Yaskawa INFORM job: UTEST.JBI

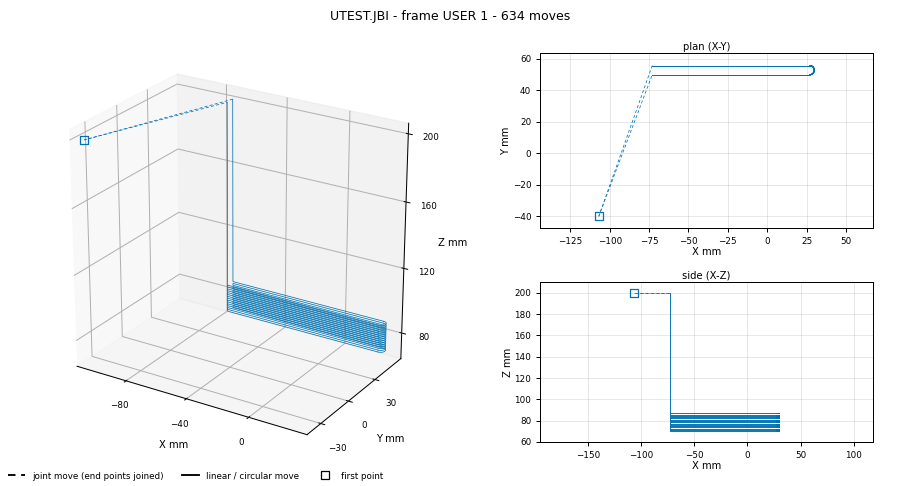
[picture p0: tool path of UTEST.JBI in frame USER 1, 634 of 649 moves have a stored position in this frame; points joined in program order, loops and branches not executed]
/JOB
//NAME UTEST
//POS
///NPOS 649,0,0,0,0,0
///USER 1
///TOOL 1
///POSTYPE USER
///RECTAN
///RCONF 1,0,0,0,0,0,0,0,0,0,0,0,0,0,0,0,0,0,0,0,0,0,0,0
C00000=-107.000,-40.000,200.000,0.0000,0.0000,-150.0000
C00001=-73.000,50.000,200.000,0.0000,0.0000,-150.0000
C00002=-73.000,50.000,70.000,0.0000,0.0000,-150.0000
C00003=-68.000,50.000,70.000,0.0000,0.0000,-150.0000
C00004=-63.000,50.000,70.000,0.0000,0.0000,-150.0000
C00005=-58.000,50.000,70.000,0.0000,0.0000,-150.0000
C00006=-53.000,50.000,70.000,0.0000,0.0000,-150.0000
C00007=-48.000,50.000,70.000,0.0000,0.0000,-150.0000
C00008=-43.000,50.000,70.000,0.0000,0.0000,-150.0000
C00009=-38.000,50.000,70.000,0.0000,0.0000,-150.0000
C00010=-33.000,50.000,70.000,0.0000,0.0000,-150.0000
C00011=-28.000,50.000,70.000,0.0000,0.0000,-150.0000
C00012=-23.000,50.000,70.000,0.0000,0.0000,-150.0000
C00013=-18.000,50.000,70.000,0.0000,0.0000,-150.0000
C00014=-13.000,50.000,70.000,0.0000,0.0000,-150.0000
C00015=-8.000,50.000,70.000,0.0000,0.0000,-150.0000
C00016=-3.000,50.000,70.000,0.0000,0.0000,-150.0000
C00017=2.000,50.000,70.000,0.0000,0.0000,-150.0000
C00018=7.000,50.000,70.000,0.0000,0.0000,-150.0000
C00019=12.000,50.000,70.000,0.0000,0.0000,-150.0000
C00020=17.000,50.000,70.000,0.0000,0.0000,-150.0000
C00021=22.000,50.000,70.000,0.0000,0.0000,-150.0000
C00022=27.000,50.000,70.000,0.0000,0.0000,-150.0000
C00023=29.915,52.915,70.000,0.0000,0.0000,-150.0000
C00024=27.000,55.829,70.000,0.0000,0.0000,-150.0000
C00025=22.000,55.829,70.000,0.0000,0.0000,-150.0000
C00026=17.000,55.829,70.000,0.0000,0.0000,-150.0000
C00027=12.000,55.829,70.000,0.0000,0.0000,-150.0000
C00028=7.000,55.829,70.000,0.0000,0.0000,-150.0000
C00029=2.000,55.829,70.000,0.0000,0.0000,-150.0000
C00030=-3.000,55.829,70.000,0.0000,0.0000,-150.0000
C00031=-8.000,55.829,70.000,0.0000,0.0000,-150.0000
C00032=-13.000,55.829,70.000,0.0000,0.0000,-150.0000
C00033=-18.000,55.829,70.000,0.0000,0.0000,-150.0000
C00034=-23.000,55.829,70.000,0.0000,0.0000,-150.0000
C00035=-28.000,55.829,70.000,0.0000,0.0000,-150.0000
C00036=-33.000,55.829,70.000,0.0000,0.0000,-150.0000
C00037=-38.000,55.829,70.000,0.0000,0.0000,-150.0000
C00038=-43.000,55.829,70.000,0.0000,0.0000,-150.0000
C00039=-48.000,55.829,70.000,0.0000,0.0000,-150.0000
C00040=-53.000,55.829,70.000,0.0000,0.0000,-150.0000
C00041=-58.000,55.829,70.000,0.0000,0.0000,-150.0000
C00042=-63.000,55.829,70.000,0.0000,0.0000,-150.0000
C00043=-68.000,55.829,70.000,0.0000,0.0000,-150.0000
C00044=-73.000,55.829,70.000,0.0000,0.0000,-150.0000
C00045=-73.000,55.829,71.200,0.0000,0.0000,-150.0000
C00046=-68.000,55.829,71.200,0.0000,0.0000,-150.0000
C00047=-63.000,55.829,71.200,0.0000,0.0000,-150.0000
C00048=-58.000,55.829,71.200,0.0000,0.0000,-150.0000
C00049=-53.000,55.829,71.200,0.0000,0.0000,-150.0000
C00050=-48.000,55.829,71.200,0.0000,0.0000,-150.0000
C00051=-43.000,55.829,71.200,0.0000,0.0000,-150.0000
C00052=-38.000,55.829,71.200,0.0000,0.0000,-150.0000
C00053=-33.000,55.829,71.200,0.0000,0.0000,-150.0000
C00054=-28.000,55.829,71.200,0.0000,0.0000,-150.0000
C00055=-23.000,55.829,71.200,0.0000,0.0000,-150.0000
C00056=-18.000,55.829,71.200,0.0000,0.0000,-150.0000
C00057=-13.000,55.829,71.200,0.0000,0.0000,-150.0000
C00058=-8.000,55.829,71.200,0.0000,0.0000,-150.0000
C00059=-3.000,55.829,71.200,0.0000,0.0000,-150.0000
C00060=2.000,55.829,71.200,0.0000,0.0000,-150.0000
C00061=7.000,55.829,71.200,0.0000,0.0000,-150.0000
C00062=12.000,55.829,71.200,0.0000,0.0000,-150.0000
C00063=17.000,55.829,71.200,0.0000,0.0000,-150.0000
C00064=22.000,55.829,71.200,0.0000,0.0000,-150.0000
C00065=27.000,55.829,71.200,0.0000,0.0000,-150.0000
C00066=29.915,52.915,71.200,0.0000,0.0000,-150.0000
C00067=27.000,50.000,71.200,0.0000,0.0000,-150.0000
C00068=22.000,50.000,71.200,0.0000,0.0000,-150.0000
C00069=17.000,50.000,71.200,0.0000,0.0000,-150.0000
C00070=12.000,50.000,71.200,0.0000,0.0000,-150.0000
C00071=7.000,50.000,71.200,0.0000,0.0000,-150.0000
C00072=2.000,50.000,71.200,0.0000,0.0000,-150.0000
C00073=-3.000,50.000,71.200,0.0000,0.0000,-150.0000
C00074=-8.000,50.000,71.200,0.0000,0.0000,-150.0000
C00075=-13.000,50.000,71.200,0.0000,0.0000,-150.0000
C00076=-18.000,50.000,71.200,0.0000,0.0000,-150.0000
C00077=-23.000,50.000,71.200,0.0000,0.0000,-150.0000
C00078=-28.000,50.000,71.200,0.0000,0.0000,-150.0000
C00079=-33.000,50.000,71.200,0.0000,0.0000,-150.0000
C00080=-38.000,50.000,71.200,0.0000,0.0000,-150.0000
C00081=-43.000,50.000,71.200,0.0000,0.0000,-150.0000
C00082=-48.000,50.000,71.200,0.0000,0.0000,-150.0000
C00083=-53.000,50.000,71.200,0.0000,0.0000,-150.0000
C00084=-58.000,50.000,71.200,0.0000,0.0000,-150.0000
C00085=-63.000,50.000,71.200,0.0000,0.0000,-150.0000
C00086=-68.000,50.000,71.200,0.0000,0.0000,-150.0000
C00087=-73.000,50.000,71.200,0.0000,0.0000,-150.0000
C00088=-73.000,50.000,72.400,0.0000,0.0000,-150.0000
C00089=-68.000,50.000,72.400,0.0000,0.0000,-150.0000
C00090=-63.000,50.000,72.400,0.0000,0.0000,-150.0000
C00091=-58.000,50.000,72.400,0.0000,0.0000,-150.0000
C00092=-53.000,50.000,72.400,0.0000,0.0000,-150.0000
C00093=-48.000,50.000,72.400,0.0000,0.0000,-150.0000
C00094=-43.000,50.000,72.400,0.0000,0.0000,-150.0000
C00095=-38.000,50.000,72.400,0.0000,0.0000,-150.0000
C00096=-33.000,50.000,72.400,0.0000,0.0000,-150.0000
C00097=-28.000,50.000,72.400,0.0000,0.0000,-150.0000
C00098=-23.000,50.000,72.400,0.0000,0.0000,-150.0000
C00099=-18.000,50.000,72.400,0.0000,0.0000,-150.0000
C00100=-13.000,50.000,72.400,0.0000,0.0000,-150.0000
C00101=-8.000,50.000,72.400,0.0000,0.0000,-150.0000
C00102=-3.000,50.000,72.400,0.0000,0.0000,-150.0000
C00103=2.000,50.000,72.400,0.0000,0.0000,-150.0000
C00104=7.000,50.000,72.400,0.0000,0.0000,-150.0000
C00105=12.000,50.000,72.400,0.0000,0.0000,-150.0000
C00106=17.000,50.000,72.400,0.0000,0.0000,-150.0000
C00107=22.000,50.000,72.400,0.0000,0.0000,-150.0000
C00108=27.000,50.000,72.400,0.0000,0.0000,-150.0000
C00109=29.915,52.915,72.400,0.0000,0.0000,-150.0000
C00110=27.000,55.829,72.400,0.0000,0.0000,-150.0000
C00111=22.000,55.829,72.400,0.0000,0.0000,-150.0000
C00112=17.000,55.829,72.400,0.0000,0.0000,-150.0000
C00113=12.000,55.829,72.400,0.0000,0.0000,-150.0000
C00114=7.000,55.829,72.400,0.0000,0.0000,-150.0000
C00115=2.000,55.829,72.400,0.0000,0.0000,-150.0000
C00116=-3.000,55.829,72.400,0.0000,0.0000,-150.0000
C00117=-8.000,55.829,72.400,0.0000,0.0000,-150.0000
C00118=-13.000,55.829,72.400,0.0000,0.0000,-150.0000
C00119=-18.000,55.829,72.400,0.0000,0.0000,-150.0000
C00120=-23.000,55.829,72.400,0.0000,0.0000,-150.0000
C00121=-28.000,55.829,72.400,0.0000,0.0000,-150.0000
C00122=-33.000,55.829,72.400,0.0000,0.0000,-150.0000
C00123=-38.000,55.829,72.400,0.0000,0.0000,-150.0000
C00124=-43.000,55.829,72.400,0.0000,0.0000,-150.0000
C00125=-48.000,55.829,72.400,0.0000,0.0000,-150.0000
C00126=-53.000,55.829,72.400,0.0000,0.0000,-150.0000
C00127=-58.000,55.829,72.400,0.0000,0.0000,-150.0000
C00128=-63.000,55.829,72.400,0.0000,0.0000,-150.0000
C00129=-68.000,55.829,72.400,0.0000,0.0000,-150.0000
C00130=-73.000,55.829,72.400,0.0000,0.0000,-150.0000
C00131=-73.000,55.829,73.600,0.0000,0.0000,-150.0000
C00132=-68.000,55.829,73.600,0.0000,0.0000,-150.0000
C00133=-63.000,55.829,73.600,0.0000,0.0000,-150.0000
C00134=-58.000,55.829,73.600,0.0000,0.0000,-150.0000
C00135=-53.000,55.829,73.600,0.0000,0.0000,-150.0000
C00136=-48.000,55.829,73.600,0.0000,0.0000,-150.0000
C00137=-43.000,55.829,73.600,0.0000,0.0000,-150.0000
C00138=-38.000,55.829,73.600,0.0000,0.0000,-150.0000
C00139=-33.000,55.829,73.600,0.0000,0.0000,-150.0000
C00140=-28.000,55.829,73.600,0.0000,0.0000,-150.0000
C00141=-23.000,55.829,73.600,0.0000,0.0000,-150.0000
C00142=-18.000,55.829,73.600,0.0000,0.0000,-150.0000
C00143=-13.000,55.829,73.600,0.0000,0.0000,-150.0000
C00144=-8.000,55.829,73.600,0.0000,0.0000,-150.0000
C00145=-3.000,55.829,73.600,0.0000,0.0000,-150.0000
C00146=2.000,55.829,73.600,0.0000,0.0000,-150.0000
C00147=7.000,55.829,73.600,0.0000,0.0000,-150.0000
C00148=12.000,55.829,73.600,0.0000,0.0000,-150.0000
C00149=17.000,55.829,73.600,0.0000,0.0000,-150.0000
C00150=22.000,55.829,73.600,0.0000,0.0000,-150.0000
C00151=27.000,55.829,73.600,0.0000,0.0000,-150.0000
C00152=29.915,52.915,73.600,0.0000,0.0000,-150.0000
C00153=27.000,50.000,73.600,0.0000,0.0000,-150.0000
C00154=22.000,50.000,73.600,0.0000,0.0000,-150.0000
C00155=17.000,50.000,73.600,0.0000,0.0000,-150.0000
C00156=12.000,50.000,73.600,0.0000,0.0000,-150.0000
C00157=7.000,50.000,73.600,0.0000,0.0000,-150.0000
C00158=2.000,50.000,73.600,0.0000,0.0000,-150.0000
C00159=-3.000,50.000,73.600,0.0000,0.0000,-150.0000
C00160=-8.000,50.000,73.600,0.0000,0.0000,-150.0000
C00161=-13.000,50.000,73.600,0.0000,0.0000,-150.0000
C00162=-18.000,50.000,73.600,0.0000,0.0000,-150.0000
C00163=-23.000,50.000,73.600,0.0000,0.0000,-150.0000
C00164=-28.000,50.000,73.600,0.0000,0.0000,-150.0000
C00165=-33.000,50.000,73.600,0.0000,0.0000,-150.0000
C00166=-38.000,50.000,73.600,0.0000,0.0000,-150.0000
C00167=-43.000,50.000,73.600,0.0000,0.0000,-150.0000
C00168=-48.000,50.000,73.600,0.0000,0.0000,-150.0000
C00169=-53.000,50.000,73.600,0.0000,0.0000,-150.0000
C00170=-58.000,50.000,73.600,0.0000,0.0000,-150.0000
C00171=-63.000,50.000,73.600,0.0000,0.0000,-150.0000
C00172=-68.000,50.000,73.600,0.0000,0.0000,-150.0000
C00173=-73.000,50.000,73.600,0.0000,0.0000,-150.0000
C00174=-73.000,50.000,74.800,0.0000,0.0000,-150.0000
C00175=-68.000,50.000,74.800,0.0000,0.0000,-150.0000
C00176=-63.000,50.000,74.800,0.0000,0.0000,-150.0000
C00177=-58.000,50.000,74.800,0.0000,0.0000,-150.0000
C00178=-53.000,50.000,74.800,0.0000,0.0000,-150.0000
C00179=-48.000,50.000,74.800,0.0000,0.0000,-150.0000
C00180=-43.000,50.000,74.800,0.0000,0.0000,-150.0000
C00181=-38.000,50.000,74.800,0.0000,0.0000,-150.0000
C00182=-33.000,50.000,74.800,0.0000,0.0000,-150.0000
C00183=-28.000,50.000,74.800,0.0000,0.0000,-150.0000
C00184=-23.000,50.000,74.800,0.0000,0.0000,-150.0000
C00185=-18.000,50.000,74.800,0.0000,0.0000,-150.0000
C00186=-13.000,50.000,74.800,0.0000,0.0000,-150.0000
C00187=-8.000,50.000,74.800,0.0000,0.0000,-150.0000
C00188=-3.000,50.000,74.800,0.0000,0.0000,-150.0000
C00189=2.000,50.000,74.800,0.0000,0.0000,-150.0000
C00190=7.000,50.000,74.800,0.0000,0.0000,-150.0000
C00191=12.000,50.000,74.800,0.0000,0.0000,-150.0000
C00192=17.000,50.000,74.800,0.0000,0.0000,-150.0000
C00193=22.000,50.000,74.800,0.0000,0.0000,-150.0000
C00194=27.000,50.000,74.800,0.0000,0.0000,-150.0000
C00195=29.915,52.915,74.800,0.0000,0.0000,-150.0000
C00196=27.000,55.829,74.800,0.0000,0.0000,-150.0000
C00197=22.000,55.829,74.800,0.0000,0.0000,-150.0000
C00198=17.000,55.829,74.800,0.0000,0.0000,-150.0000
C00199=12.000,55.829,74.800,0.0000,0.0000,-150.0000
C00200=7.000,55.829,74.800,0.0000,0.0000,-150.0000
C00201=2.000,55.829,74.800,0.0000,0.0000,-150.0000
C00202=-3.000,55.829,74.800,0.0000,0.0000,-150.0000
C00203=-8.000,55.829,74.800,0.0000,0.0000,-150.0000
C00204=-13.000,55.829,74.800,0.0000,0.0000,-150.0000
C00205=-18.000,55.829,74.800,0.0000,0.0000,-150.0000
C00206=-23.000,55.829,74.800,0.0000,0.0000,-150.0000
C00207=-28.000,55.829,74.800,0.0000,0.0000,-150.0000
C00208=-33.000,55.829,74.800,0.0000,0.0000,-150.0000
C00209=-38.000,55.829,74.800,0.0000,0.0000,-150.0000
C00210=-43.000,55.829,74.800,0.0000,0.0000,-150.0000
C00211=-48.000,55.829,74.800,0.0000,0.0000,-150.0000
C00212=-53.000,55.829,74.800,0.0000,0.0000,-150.0000
C00213=-58.000,55.829,74.800,0.0000,0.0000,-150.0000
C00214=-63.000,55.829,74.800,0.0000,0.0000,-150.0000
C00215=-68.000,55.829,74.800,0.0000,0.0000,-150.0000
C00216=-73.000,55.829,74.800,0.0000,0.0000,-150.0000
C00217=-73.000,55.829,76.000,0.0000,0.0000,-150.0000
C00218=-68.000,55.829,76.000,0.0000,0.0000,-150.0000
C00219=-63.000,55.829,76.000,0.0000,0.0000,-150.0000
C00220=-58.000,55.829,76.000,0.0000,0.0000,-150.0000
C00221=-53.000,55.829,76.000,0.0000,0.0000,-150.0000
C00222=-48.000,55.829,76.000,0.0000,0.0000,-150.0000
C00223=-43.000,55.829,76.000,0.0000,0.0000,-150.0000
C00224=-38.000,55.829,76.000,0.0000,0.0000,-150.0000
C00225=-33.000,55.829,76.000,0.0000,0.0000,-150.0000
C00226=-28.000,55.829,76.000,0.0000,0.0000,-150.0000
C00227=-23.000,55.829,76.000,0.0000,0.0000,-150.0000
C00228=-18.000,55.829,76.000,0.0000,0.0000,-150.0000
C00229=-13.000,55.829,76.000,0.0000,0.0000,-150.0000
C00230=-8.000,55.829,76.000,0.0000,0.0000,-150.0000
C00231=-3.000,55.829,76.000,0.0000,0.0000,-150.0000
C00232=2.000,55.829,76.000,0.0000,0.0000,-150.0000
C00233=7.000,55.829,76.000,0.0000,0.0000,-150.0000
C00234=12.000,55.829,76.000,0.0000,0.0000,-150.0000
C00235=17.000,55.829,76.000,0.0000,0.0000,-150.0000
C00236=22.000,55.829,76.000,0.0000,0.0000,-150.0000
C00237=27.000,55.829,76.000,0.0000,0.0000,-150.0000
C00238=29.915,52.915,76.000,0.0000,0.0000,-150.0000
C00239=27.000,50.000,76.000,0.0000,0.0000,-150.0000
C00240=22.000,50.000,76.000,0.0000,0.0000,-150.0000
C00241=17.000,50.000,76.000,0.0000,0.0000,-150.0000
C00242=12.000,50.000,76.000,0.0000,0.0000,-150.0000
C00243=7.000,50.000,76.000,0.0000,0.0000,-150.0000
C00244=2.000,50.000,76.000,0.0000,0.0000,-150.0000
C00245=-3.000,50.000,76.000,0.0000,0.0000,-150.0000
C00246=-8.000,50.000,76.000,0.0000,0.0000,-150.0000
C00247=-13.000,50.000,76.000,0.0000,0.0000,-150.0000
C00248=-18.000,50.000,76.000,0.0000,0.0000,-150.0000
C00249=-23.000,50.000,76.000,0.0000,0.0000,-150.0000
C00250=-28.000,50.000,76.000,0.0000,0.0000,-150.0000
C00251=-33.000,50.000,76.000,0.0000,0.0000,-150.0000
C00252=-38.000,50.000,76.000,0.0000,0.0000,-150.0000
C00253=-43.000,50.000,76.000,0.0000,0.0000,-150.0000
C00254=-48.000,50.000,76.000,0.0000,0.0000,-150.0000
C00255=-53.000,50.000,76.000,0.0000,0.0000,-150.0000
C00256=-58.000,50.000,76.000,0.0000,0.0000,-150.0000
C00257=-63.000,50.000,76.000,0.0000,0.0000,-150.0000
C00258=-68.000,50.000,76.000,0.0000,0.0000,-150.0000
C00259=-73.000,50.000,76.000,0.0000,0.0000,-150.0000
C00260=-73.000,50.000,77.200,0.0000,0.0000,-150.0000
C00261=-68.000,50.000,77.200,0.0000,0.0000,-150.0000
C00262=-63.000,50.000,77.200,0.0000,0.0000,-150.0000
C00263=-58.000,50.000,77.200,0.0000,0.0000,-150.0000
C00264=-53.000,50.000,77.200,0.0000,0.0000,-150.0000
C00265=-48.000,50.000,77.200,0.0000,0.0000,-150.0000
C00266=-43.000,50.000,77.200,0.0000,0.0000,-150.0000
C00267=-38.000,50.000,77.200,0.0000,0.0000,-150.0000
C00268=-33.000,50.000,77.200,0.0000,0.0000,-150.0000
C00269=-28.000,50.000,77.200,0.0000,0.0000,-150.0000
C00270=-23.000,50.000,77.200,0.0000,0.0000,-150.0000
C00271=-18.000,50.000,77.200,0.0000,0.0000,-150.0000
C00272=-13.000,50.000,77.200,0.0000,0.0000,-150.0000
C00273=-8.000,50.000,77.200,0.0000,0.0000,-150.0000
C00274=-3.000,50.000,77.200,0.0000,0.0000,-150.0000
C00275=2.000,50.000,77.200,0.0000,0.0000,-150.0000
C00276=7.000,50.000,77.200,0.0000,0.0000,-150.0000
C00277=12.000,50.000,77.200,0.0000,0.0000,-150.0000
C00278=17.000,50.000,77.200,0.0000,0.0000,-150.0000
C00279=22.000,50.000,77.200,0.0000,0.0000,-150.0000
C00280=27.000,50.000,77.200,0.0000,0.0000,-150.0000
C00281=29.915,52.915,77.200,0.0000,0.0000,-150.0000
C00282=27.000,55.829,77.200,0.0000,0.0000,-150.0000
C00283=22.000,55.829,77.200,0.0000,0.0000,-150.0000
C00284=17.000,55.829,77.200,0.0000,0.0000,-150.0000
C00285=12.000,55.829,77.200,0.0000,0.0000,-150.0000
C00286=7.000,55.829,77.200,0.0000,0.0000,-150.0000
C00287=2.000,55.829,77.200,0.0000,0.0000,-150.0000
C00288=-3.000,55.829,77.200,0.0000,0.0000,-150.0000
C00289=-8.000,55.829,77.200,0.0000,0.0000,-150.0000
C00290=-13.000,55.829,77.200,0.0000,0.0000,-150.0000
C00291=-18.000,55.829,77.200,0.0000,0.0000,-150.0000
C00292=-23.000,55.829,77.200,0.0000,0.0000,-150.0000
C00293=-28.000,55.829,77.200,0.0000,0.0000,-150.0000
C00294=-33.000,55.829,77.200,0.0000,0.0000,-150.0000
C00295=-38.000,55.829,77.200,0.0000,0.0000,-150.0000
C00296=-43.000,55.829,77.200,0.0000,0.0000,-150.0000
C00297=-48.000,55.829,77.200,0.0000,0.0000,-150.0000
C00298=-53.000,55.829,77.200,0.0000,0.0000,-150.0000
C00299=-58.000,55.829,77.200,0.0000,0.0000,-150.0000
C00300=-63.000,55.829,77.200,0.0000,0.0000,-150.0000
C00301=-68.000,55.829,77.200,0.0000,0.0000,-150.0000
C00302=-73.000,55.829,77.200,0.0000,0.0000,-150.0000
C00303=-73.000,55.829,78.400,0.0000,0.0000,-150.0000
C00304=-68.000,55.829,78.400,0.0000,0.0000,-150.0000
C00305=-63.000,55.829,78.400,0.0000,0.0000,-150.0000
C00306=-58.000,55.829,78.400,0.0000,0.0000,-150.0000
C00307=-53.000,55.829,78.400,0.0000,0.0000,-150.0000
C00308=-48.000,55.829,78.400,0.0000,0.0000,-150.0000
C00309=-43.000,55.829,78.400,0.0000,0.0000,-150.0000
C00310=-38.000,55.829,78.400,0.0000,0.0000,-150.0000
C00311=-33.000,55.829,78.400,0.0000,0.0000,-150.0000
C00312=-28.000,55.829,78.400,0.0000,0.0000,-150.0000
C00313=-23.000,55.829,78.400,0.0000,0.0000,-150.0000
C00314=-18.000,55.829,78.400,0.0000,0.0000,-150.0000
C00315=-13.000,55.829,78.400,0.0000,0.0000,-150.0000
C00316=-8.000,55.829,78.400,0.0000,0.0000,-150.0000
C00317=-3.000,55.829,78.400,0.0000,0.0000,-150.0000
C00318=2.000,55.829,78.400,0.0000,0.0000,-150.0000
C00319=7.000,55.829,78.400,0.0000,0.0000,-150.0000
C00320=12.000,55.829,78.400,0.0000,0.0000,-150.0000
C00321=17.000,55.829,78.400,0.0000,0.0000,-150.0000
C00322=22.000,55.829,78.400,0.0000,0.0000,-150.0000
C00323=27.000,55.829,78.400,0.0000,0.0000,-150.0000
C00324=29.915,52.915,78.400,0.0000,0.0000,-150.0000
C00325=27.000,50.000,78.400,0.0000,0.0000,-150.0000
C00326=22.000,50.000,78.400,0.0000,0.0000,-150.0000
C00327=17.000,50.000,78.400,0.0000,0.0000,-150.0000
C00328=12.000,50.000,78.400,0.0000,0.0000,-150.0000
C00329=7.000,50.000,78.400,0.0000,0.0000,-150.0000
C00330=2.000,50.000,78.400,0.0000,0.0000,-150.0000
C00331=-3.000,50.000,78.400,0.0000,0.0000,-150.0000
C00332=-8.000,50.000,78.400,0.0000,0.0000,-150.0000
C00333=-13.000,50.000,78.400,0.0000,0.0000,-150.0000
C00334=-18.000,50.000,78.400,0.0000,0.0000,-150.0000
C00335=-23.000,50.000,78.400,0.0000,0.0000,-150.0000
C00336=-28.000,50.000,78.400,0.0000,0.0000,-150.0000
C00337=-33.000,50.000,78.400,0.0000,0.0000,-150.0000
C00338=-38.000,50.000,78.400,0.0000,0.0000,-150.0000
C00339=-43.000,50.000,78.400,0.0000,0.0000,-150.0000
C00340=-48.000,50.000,78.400,0.0000,0.0000,-150.0000
C00341=-53.000,50.000,78.400,0.0000,0.0000,-150.0000
C00342=-58.000,50.000,78.400,0.0000,0.0000,-150.0000
C00343=-63.000,50.000,78.400,0.0000,0.0000,-150.0000
C00344=-68.000,50.000,78.400,0.0000,0.0000,-150.0000
C00345=-73.000,50.000,78.400,0.0000,0.0000,-150.0000
C00346=-73.000,50.000,79.600,0.0000,0.0000,-150.0000
C00347=-68.000,50.000,79.600,0.0000,0.0000,-150.0000
C00348=-63.000,50.000,79.600,0.0000,0.0000,-150.0000
C00349=-58.000,50.000,79.600,0.0000,0.0000,-150.0000
C00350=-53.000,50.000,79.600,0.0000,0.0000,-150.0000
C00351=-48.000,50.000,79.600,0.0000,0.0000,-150.0000
C00352=-43.000,50.000,79.600,0.0000,0.0000,-150.0000
C00353=-38.000,50.000,79.600,0.0000,0.0000,-150.0000
C00354=-33.000,50.000,79.600,0.0000,0.0000,-150.0000
C00355=-28.000,50.000,79.600,0.0000,0.0000,-150.0000
C00356=-23.000,50.000,79.600,0.0000,0.0000,-150.0000
C00357=-18.000,50.000,79.600,0.0000,0.0000,-150.0000
C00358=-13.000,50.000,79.600,0.0000,0.0000,-150.0000
C00359=-8.000,50.000,79.600,0.0000,0.0000,-150.0000
C00360=-3.000,50.000,79.600,0.0000,0.0000,-150.0000
C00361=2.000,50.000,79.600,0.0000,0.0000,-150.0000
C00362=7.000,50.000,79.600,0.0000,0.0000,-150.0000
C00363=12.000,50.000,79.600,0.0000,0.0000,-150.0000
C00364=17.000,50.000,79.600,0.0000,0.0000,-150.0000
C00365=22.000,50.000,79.600,0.0000,0.0000,-150.0000
C00366=27.000,50.000,79.600,0.0000,0.0000,-150.0000
C00367=29.915,52.915,79.600,0.0000,0.0000,-150.0000
C00368=27.000,55.829,79.600,0.0000,0.0000,-150.0000
C00369=22.000,55.829,79.600,0.0000,0.0000,-150.0000
C00370=17.000,55.829,79.600,0.0000,0.0000,-150.0000
C00371=12.000,55.829,79.600,0.0000,0.0000,-150.0000
C00372=7.000,55.829,79.600,0.0000,0.0000,-150.0000
C00373=2.000,55.829,79.600,0.0000,0.0000,-150.0000
C00374=-3.000,55.829,79.600,0.0000,0.0000,-150.0000
C00375=-8.000,55.829,79.600,0.0000,0.0000,-150.0000
C00376=-13.000,55.829,79.600,0.0000,0.0000,-150.0000
C00377=-18.000,55.829,79.600,0.0000,0.0000,-150.0000
C00378=-23.000,55.829,79.600,0.0000,0.0000,-150.0000
C00379=-28.000,55.829,79.600,0.0000,0.0000,-150.0000
C00380=-33.000,55.829,79.600,0.0000,0.0000,-150.0000
C00381=-38.000,55.829,79.600,0.0000,0.0000,-150.0000
C00382=-43.000,55.829,79.600,0.0000,0.0000,-150.0000
C00383=-48.000,55.829,79.600,0.0000,0.0000,-150.0000
C00384=-53.000,55.829,79.600,0.0000,0.0000,-150.0000
C00385=-58.000,55.829,79.600,0.0000,0.0000,-150.0000
C00386=-63.000,55.829,79.600,0.0000,0.0000,-150.0000
C00387=-68.000,55.829,79.600,0.0000,0.0000,-150.0000
C00388=-73.000,55.829,79.600,0.0000,0.0000,-150.0000
C00389=-73.000,55.829,80.800,0.0000,0.0000,-150.0000
C00390=-68.000,55.829,80.800,0.0000,0.0000,-150.0000
C00391=-63.000,55.829,80.800,0.0000,0.0000,-150.0000
C00392=-58.000,55.829,80.800,0.0000,0.0000,-150.0000
C00393=-53.000,55.829,80.800,0.0000,0.0000,-150.0000
C00394=-48.000,55.829,80.800,0.0000,0.0000,-150.0000
C00395=-43.000,55.829,80.800,0.0000,0.0000,-150.0000
C00396=-38.000,55.829,80.800,0.0000,0.0000,-150.0000
C00397=-33.000,55.829,80.800,0.0000,0.0000,-150.0000
C00398=-28.000,55.829,80.800,0.0000,0.0000,-150.0000
C00399=-23.000,55.829,80.800,0.0000,0.0000,-150.0000
C00400=-18.000,55.829,80.800,0.0000,0.0000,-150.0000
C00401=-13.000,55.829,80.800,0.0000,0.0000,-150.0000
C00402=-8.000,55.829,80.800,0.0000,0.0000,-150.0000
C00403=-3.000,55.829,80.800,0.0000,0.0000,-150.0000
C00404=2.000,55.829,80.800,0.0000,0.0000,-150.0000
C00405=7.000,55.829,80.800,0.0000,0.0000,-150.0000
C00406=12.000,55.829,80.800,0.0000,0.0000,-150.0000
C00407=17.000,55.829,80.800,0.0000,0.0000,-150.0000
C00408=22.000,55.829,80.800,0.0000,0.0000,-150.0000
C00409=27.000,55.829,80.800,0.0000,0.0000,-150.0000
C00410=29.915,52.915,80.800,0.0000,0.0000,-150.0000
C00411=27.000,50.000,80.800,0.0000,0.0000,-150.0000
C00412=22.000,50.000,80.800,0.0000,0.0000,-150.0000
C00413=17.000,50.000,80.800,0.0000,0.0000,-150.0000
C00414=12.000,50.000,80.800,0.0000,0.0000,-150.0000
C00415=7.000,50.000,80.800,0.0000,0.0000,-150.0000
C00416=2.000,50.000,80.800,0.0000,0.0000,-150.0000
C00417=-3.000,50.000,80.800,0.0000,0.0000,-150.0000
C00418=-8.000,50.000,80.800,0.0000,0.0000,-150.0000
C00419=-13.000,50.000,80.800,0.0000,0.0000,-150.0000
C00420=-18.000,50.000,80.800,0.0000,0.0000,-150.0000
C00421=-23.000,50.000,80.800,0.0000,0.0000,-150.0000
C00422=-28.000,50.000,80.800,0.0000,0.0000,-150.0000
C00423=-33.000,50.000,80.800,0.0000,0.0000,-150.0000
C00424=-38.000,50.000,80.800,0.0000,0.0000,-150.0000
C00425=-43.000,50.000,80.800,0.0000,0.0000,-150.0000
C00426=-48.000,50.000,80.800,0.0000,0.0000,-150.0000
C00427=-53.000,50.000,80.800,0.0000,0.0000,-150.0000
C00428=-58.000,50.000,80.800,0.0000,0.0000,-150.0000
C00429=-63.000,50.000,80.800,0.0000,0.0000,-150.0000
C00430=-68.000,50.000,80.800,0.0000,0.0000,-150.0000
C00431=-73.000,50.000,80.800,0.0000,0.0000,-150.0000
C00432=-73.000,50.000,82.000,0.0000,0.0000,-150.0000
C00433=-68.000,50.000,82.000,0.0000,0.0000,-150.0000
C00434=-63.000,50.000,82.000,0.0000,0.0000,-150.0000
C00435=-58.000,50.000,82.000,0.0000,0.0000,-150.0000
C00436=-53.000,50.000,82.000,0.0000,0.0000,-150.0000
C00437=-48.000,50.000,82.000,0.0000,0.0000,-150.0000
C00438=-43.000,50.000,82.000,0.0000,0.0000,-150.0000
C00439=-38.000,50.000,82.000,0.0000,0.0000,-150.0000
C00440=-33.000,50.000,82.000,0.0000,0.0000,-150.0000
C00441=-28.000,50.000,82.000,0.0000,0.0000,-150.0000
C00442=-23.000,50.000,82.000,0.0000,0.0000,-150.0000
C00443=-18.000,50.000,82.000,0.0000,0.0000,-150.0000
C00444=-13.000,50.000,82.000,0.0000,0.0000,-150.0000
C00445=-8.000,50.000,82.000,0.0000,0.0000,-150.0000
C00446=-3.000,50.000,82.000,0.0000,0.0000,-150.0000
C00447=2.000,50.000,82.000,0.0000,0.0000,-150.0000
C00448=7.000,50.000,82.000,0.0000,0.0000,-150.0000
C00449=12.000,50.000,82.000,0.0000,0.0000,-150.0000
C00450=17.000,50.000,82.000,0.0000,0.0000,-150.0000
C00451=22.000,50.000,82.000,0.0000,0.0000,-150.0000
C00452=27.000,50.000,82.000,0.0000,0.0000,-150.0000
C00453=29.915,52.915,82.000,0.0000,0.0000,-150.0000
C00454=27.000,55.829,82.000,0.0000,0.0000,-150.0000
C00455=22.000,55.829,82.000,0.0000,0.0000,-150.0000
C00456=17.000,55.829,82.000,0.0000,0.0000,-150.0000
C00457=12.000,55.829,82.000,0.0000,0.0000,-150.0000
C00458=7.000,55.829,82.000,0.0000,0.0000,-150.0000
C00459=2.000,55.829,82.000,0.0000,0.0000,-150.0000
C00460=-3.000,55.829,82.000,0.0000,0.0000,-150.0000
C00461=-8.000,55.829,82.000,0.0000,0.0000,-150.0000
C00462=-13.000,55.829,82.000,0.0000,0.0000,-150.0000
C00463=-18.000,55.829,82.000,0.0000,0.0000,-150.0000
C00464=-23.000,55.829,82.000,0.0000,0.0000,-150.0000
C00465=-28.000,55.829,82.000,0.0000,0.0000,-150.0000
C00466=-33.000,55.829,82.000,0.0000,0.0000,-150.0000
C00467=-38.000,55.829,82.000,0.0000,0.0000,-150.0000
C00468=-43.000,55.829,82.000,0.0000,0.0000,-150.0000
C00469=-48.000,55.829,82.000,0.0000,0.0000,-150.0000
C00470=-53.000,55.829,82.000,0.0000,0.0000,-150.0000
C00471=-58.000,55.829,82.000,0.0000,0.0000,-150.0000
C00472=-63.000,55.829,82.000,0.0000,0.0000,-150.0000
C00473=-68.000,55.829,82.000,0.0000,0.0000,-150.0000
C00474=-73.000,55.829,82.000,0.0000,0.0000,-150.0000
C00475=-73.000,55.829,83.200,0.0000,0.0000,-150.0000
C00476=-68.000,55.829,83.200,0.0000,0.0000,-150.0000
C00477=-63.000,55.829,83.200,0.0000,0.0000,-150.0000
C00478=-58.000,55.829,83.200,0.0000,0.0000,-150.0000
C00479=-53.000,55.829,83.200,0.0000,0.0000,-150.0000
C00480=-48.000,55.829,83.200,0.0000,0.0000,-150.0000
C00481=-43.000,55.829,83.200,0.0000,0.0000,-150.0000
C00482=-38.000,55.829,83.200,0.0000,0.0000,-150.0000
C00483=-33.000,55.829,83.200,0.0000,0.0000,-150.0000
C00484=-28.000,55.829,83.200,0.0000,0.0000,-150.0000
C00485=-23.000,55.829,83.200,0.0000,0.0000,-150.0000
C00486=-18.000,55.829,83.200,0.0000,0.0000,-150.0000
C00487=-13.000,55.829,83.200,0.0000,0.0000,-150.0000
C00488=-8.000,55.829,83.200,0.0000,0.0000,-150.0000
C00489=-3.000,55.829,83.200,0.0000,0.0000,-150.0000
C00490=2.000,55.829,83.200,0.0000,0.0000,-150.0000
C00491=7.000,55.829,83.200,0.0000,0.0000,-150.0000
C00492=12.000,55.829,83.200,0.0000,0.0000,-150.0000
C00493=17.000,55.829,83.200,0.0000,0.0000,-150.0000
C00494=22.000,55.829,83.200,0.0000,0.0000,-150.0000
C00495=27.000,55.829,83.200,0.0000,0.0000,-150.0000
C00496=29.915,52.915,83.200,0.0000,0.0000,-150.0000
C00497=27.000,50.000,83.200,0.0000,0.0000,-150.0000
C00498=22.000,50.000,83.200,0.0000,0.0000,-150.0000
C00499=17.000,50.000,83.200,0.0000,0.0000,-150.0000
C00500=12.000,50.000,83.200,0.0000,0.0000,-150.0000
C00501=7.000,50.000,83.200,0.0000,0.0000,-150.0000
C00502=2.000,50.000,83.200,0.0000,0.0000,-150.0000
C00503=-3.000,50.000,83.200,0.0000,0.0000,-150.0000
C00504=-8.000,50.000,83.200,0.0000,0.0000,-150.0000
C00505=-13.000,50.000,83.200,0.0000,0.0000,-150.0000
C00506=-18.000,50.000,83.200,0.0000,0.0000,-150.0000
C00507=-23.000,50.000,83.200,0.0000,0.0000,-150.0000
C00508=-28.000,50.000,83.200,0.0000,0.0000,-150.0000
C00509=-33.000,50.000,83.200,0.0000,0.0000,-150.0000
C00510=-38.000,50.000,83.200,0.0000,0.0000,-150.0000
C00511=-43.000,50.000,83.200,0.0000,0.0000,-150.0000
C00512=-48.000,50.000,83.200,0.0000,0.0000,-150.0000
C00513=-53.000,50.000,83.200,0.0000,0.0000,-150.0000
C00514=-58.000,50.000,83.200,0.0000,0.0000,-150.0000
C00515=-63.000,50.000,83.200,0.0000,0.0000,-150.0000
C00516=-68.000,50.000,83.200,0.0000,0.0000,-150.0000
C00517=-73.000,50.000,83.200,0.0000,0.0000,-150.0000
C00518=-73.000,50.000,84.400,0.0000,0.0000,-150.0000
C00519=-68.000,50.000,84.400,0.0000,0.0000,-150.0000
C00520=-63.000,50.000,84.400,0.0000,0.0000,-150.0000
C00521=-58.000,50.000,84.400,0.0000,0.0000,-150.0000
C00522=-53.000,50.000,84.400,0.0000,0.0000,-150.0000
C00523=-48.000,50.000,84.400,0.0000,0.0000,-150.0000
C00524=-43.000,50.000,84.400,0.0000,0.0000,-150.0000
C00525=-38.000,50.000,84.400,0.0000,0.0000,-150.0000
C00526=-33.000,50.000,84.400,0.0000,0.0000,-150.0000
C00527=-28.000,50.000,84.400,0.0000,0.0000,-150.0000
C00528=-23.000,50.000,84.400,0.0000,0.0000,-150.0000
C00529=-18.000,50.000,84.400,0.0000,0.0000,-150.0000
C00530=-13.000,50.000,84.400,0.0000,0.0000,-150.0000
C00531=-8.000,50.000,84.400,0.0000,0.0000,-150.0000
C00532=-3.000,50.000,84.400,0.0000,0.0000,-150.0000
C00533=2.000,50.000,84.400,0.0000,0.0000,-150.0000
C00534=7.000,50.000,84.400,0.0000,0.0000,-150.0000
C00535=12.000,50.000,84.400,0.0000,0.0000,-150.0000
C00536=17.000,50.000,84.400,0.0000,0.0000,-150.0000
C00537=22.000,50.000,84.400,0.0000,0.0000,-150.0000
C00538=27.000,50.000,84.400,0.0000,0.0000,-150.0000
C00539=29.915,52.915,84.400,0.0000,0.0000,-150.0000
C00540=27.000,55.829,84.400,0.0000,0.0000,-150.0000
C00541=22.000,55.829,84.400,0.0000,0.0000,-150.0000
C00542=17.000,55.829,84.400,0.0000,0.0000,-150.0000
C00543=12.000,55.829,84.400,0.0000,0.0000,-150.0000
C00544=7.000,55.829,84.400,0.0000,0.0000,-150.0000
C00545=2.000,55.829,84.400,0.0000,0.0000,-150.0000
C00546=-3.000,55.829,84.400,0.0000,0.0000,-150.0000
C00547=-8.000,55.829,84.400,0.0000,0.0000,-150.0000
C00548=-13.000,55.829,84.400,0.0000,0.0000,-150.0000
C00549=-18.000,55.829,84.400,0.0000,0.0000,-150.0000
C00550=-23.000,55.829,84.400,0.0000,0.0000,-150.0000
C00551=-28.000,55.829,84.400,0.0000,0.0000,-150.0000
C00552=-33.000,55.829,84.400,0.0000,0.0000,-150.0000
C00553=-38.000,55.829,84.400,0.0000,0.0000,-150.0000
C00554=-43.000,55.829,84.400,0.0000,0.0000,-150.0000
C00555=-48.000,55.829,84.400,0.0000,0.0000,-150.0000
C00556=-53.000,55.829,84.400,0.0000,0.0000,-150.0000
C00557=-58.000,55.829,84.400,0.0000,0.0000,-150.0000
C00558=-63.000,55.829,84.400,0.0000,0.0000,-150.0000
C00559=-68.000,55.829,84.400,0.0000,0.0000,-150.0000
C00560=-73.000,55.829,84.400,0.0000,0.0000,-150.0000
C00561=-73.000,55.829,85.600,0.0000,0.0000,-150.0000
C00562=-68.000,55.829,85.600,0.0000,0.0000,-150.0000
C00563=-63.000,55.829,85.600,0.0000,0.0000,-150.0000
C00564=-58.000,55.829,85.600,0.0000,0.0000,-150.0000
C00565=-53.000,55.829,85.600,0.0000,0.0000,-150.0000
C00566=-48.000,55.829,85.600,0.0000,0.0000,-150.0000
C00567=-43.000,55.829,85.600,0.0000,0.0000,-150.0000
C00568=-38.000,55.829,85.600,0.0000,0.0000,-150.0000
C00569=-33.000,55.829,85.600,0.0000,0.0000,-150.0000
C00570=-28.000,55.829,85.600,0.0000,0.0000,-150.0000
C00571=-23.000,55.829,85.600,0.0000,0.0000,-150.0000
C00572=-18.000,55.829,85.600,0.0000,0.0000,-150.0000
C00573=-13.000,55.829,85.600,0.0000,0.0000,-150.0000
C00574=-8.000,55.829,85.600,0.0000,0.0000,-150.0000
C00575=-3.000,55.829,85.600,0.0000,0.0000,-150.0000
C00576=2.000,55.829,85.600,0.0000,0.0000,-150.0000
C00577=7.000,55.829,85.600,0.0000,0.0000,-150.0000
C00578=12.000,55.829,85.600,0.0000,0.0000,-150.0000
C00579=17.000,55.829,85.600,0.0000,0.0000,-150.0000
C00580=22.000,55.829,85.600,0.0000,0.0000,-150.0000
C00581=27.000,55.829,85.600,0.0000,0.0000,-150.0000
C00582=29.915,52.915,85.600,0.0000,0.0000,-150.0000
C00583=27.000,50.000,85.600,0.0000,0.0000,-150.0000
C00584=22.000,50.000,85.600,0.0000,0.0000,-150.0000
C00585=17.000,50.000,85.600,0.0000,0.0000,-150.0000
C00586=12.000,50.000,85.600,0.0000,0.0000,-150.0000
C00587=7.000,50.000,85.600,0.0000,0.0000,-150.0000
C00588=2.000,50.000,85.600,0.0000,0.0000,-150.0000
C00589=-3.000,50.000,85.600,0.0000,0.0000,-150.0000
C00590=-8.000,50.000,85.600,0.0000,0.0000,-150.0000
C00591=-13.000,50.000,85.600,0.0000,0.0000,-150.0000
C00592=-18.000,50.000,85.600,0.0000,0.0000,-150.0000
C00593=-23.000,50.000,85.600,0.0000,0.0000,-150.0000
C00594=-28.000,50.000,85.600,0.0000,0.0000,-150.0000
C00595=-33.000,50.000,85.600,0.0000,0.0000,-150.0000
C00596=-38.000,50.000,85.600,0.0000,0.0000,-150.0000
C00597=-43.000,50.000,85.600,0.0000,0.0000,-150.0000
C00598=-48.000,50.000,85.600,0.0000,0.0000,-150.0000
C00599=-53.000,50.000,85.600,0.0000,0.0000,-150.0000
C00600=-58.000,50.000,85.600,0.0000,0.0000,-150.0000
C00601=-63.000,50.000,85.600,0.0000,0.0000,-150.0000
C00602=-68.000,50.000,85.600,0.0000,0.0000,-150.0000
C00603=-73.000,50.000,85.600,0.0000,0.0000,-150.0000
C00604=-73.000,50.000,86.800,0.0000,0.0000,-150.0000
C00605=-68.000,50.000,86.800,0.0000,0.0000,-150.0000
C00606=-63.000,50.000,86.800,0.0000,0.0000,-150.0000
C00607=-58.000,50.000,86.800,0.0000,0.0000,-150.0000
C00608=-53.000,50.000,86.800,0.0000,0.0000,-150.0000
C00609=-48.000,50.000,86.800,0.0000,0.0000,-150.0000
C00610=-43.000,50.000,86.800,0.0000,0.0000,-150.0000
C00611=-38.000,50.000,86.800,0.0000,0.0000,-150.0000
C00612=-33.000,50.000,86.800,0.0000,0.0000,-150.0000
C00613=-28.000,50.000,86.800,0.0000,0.0000,-150.0000
C00614=-23.000,50.000,86.800,0.0000,0.0000,-150.0000
C00615=-18.000,50.000,86.800,0.0000,0.0000,-150.0000
C00616=-13.000,50.000,86.800,0.0000,0.0000,-150.0000
C00617=-8.000,50.000,86.800,0.0000,0.0000,-150.0000
C00618=-3.000,50.000,86.800,0.0000,0.0000,-150.0000
C00619=2.000,50.000,86.800,0.0000,0.0000,-150.0000
C00620=7.000,50.000,86.800,0.0000,0.0000,-150.0000
C00621=12.000,50.000,86.800,0.0000,0.0000,-150.0000
C00622=17.000,50.000,86.800,0.0000,0.0000,-150.0000
C00623=22.000,50.000,86.800,0.0000,0.0000,-150.0000
C00624=27.000,50.000,86.800,0.0000,0.0000,-150.0000
C00625=29.915,52.915,86.800,0.0000,0.0000,-150.0000
C00626=27.000,55.829,86.800,0.0000,0.0000,-150.0000
C00627=22.000,55.829,86.800,0.0000,0.0000,-150.0000
C00628=17.000,55.829,86.800,0.0000,0.0000,-150.0000
C00629=12.000,55.829,86.800,0.0000,0.0000,-150.0000
C00630=7.000,55.829,86.800,0.0000,0.0000,-150.0000
C00631=2.000,55.829,86.800,0.0000,0.0000,-150.0000
C00632=-3.000,55.829,86.800,0.0000,0.0000,-150.0000
C00633=-8.000,55.829,86.800,0.0000,0.0000,-150.0000
C00634=-13.000,55.829,86.800,0.0000,0.0000,-150.0000
C00635=-18.000,55.829,86.800,0.0000,0.0000,-150.0000
C00636=-23.000,55.829,86.800,0.0000,0.0000,-150.0000
C00637=-28.000,55.829,86.800,0.0000,0.0000,-150.0000
C00638=-33.000,55.829,86.800,0.0000,0.0000,-150.0000
C00639=-38.000,55.829,86.800,0.0000,0.0000,-150.0000
C00640=-43.000,55.829,86.800,0.0000,0.0000,-150.0000
C00641=-48.000,55.829,86.800,0.0000,0.0000,-150.0000
C00642=-53.000,55.829,86.800,0.0000,0.0000,-150.0000
C00643=-58.000,55.829,86.800,0.0000,0.0000,-150.0000
C00644=-63.000,55.829,86.800,0.0000,0.0000,-150.0000
C00645=-68.000,55.829,86.800,0.0000,0.0000,-150.0000
C00646=-73.000,55.829,86.800,0.0000,0.0000,-150.0000
C00647=-73.000,55.829,200.000,0.0000,0.0000,-150.0000
C00648=-107.000,-40.000,200.000,0.0000,0.0000,-150.0000
//INST
///DATE 2026/11/25 17:59
///ATTR SC,RW,RJ
////FRAME USER 1
///GROUP1 RB1
NOP
MOVJ C00000 VJ=0.78
MOVJ C00001 VJ=0.78
MOVL C00002 V=11.0 ACC=20 DEC=20
*LAG1
MACRO1 MJ#(0) ARGF1
ARCON
MOVL C00003 V=10.0 ACC=20 DEC=20
MOVL C00004 V=10.0 ACC=20 DEC=20
MOVL C00005 V=10.0 ACC=20 DEC=20
MOVL C00006 V=10.0 ACC=20 DEC=20
MOVL C00007 V=10.0 ACC=20 DEC=20
MOVL C00008 V=10.0 ACC=20 DEC=20
MOVL C00009 V=10.0 ACC=20 DEC=20
MOVL C00010 V=10.0 ACC=20 DEC=20
MOVL C00011 V=10.0 ACC=20 DEC=20
MOVL C00012 V=10.0 ACC=20 DEC=20
MOVL C00013 V=10.0 ACC=20 DEC=20
MOVL C00014 V=10.0 ACC=20 DEC=20
MOVL C00015 V=10.0 ACC=20 DEC=20
MOVL C00016 V=10.0 ACC=20 DEC=20
MOVL C00017 V=10.0 ACC=20 DEC=20
MOVL C00018 V=10.0 ACC=20 DEC=20
MOVL C00019 V=10.0 ACC=20 DEC=20
MOVL C00020 V=10.0 ACC=20 DEC=20
MOVL C00021 V=10.0 ACC=20 DEC=20
MOVC C00022 V=14.0 ACC=20 DEC=20
MOVC C00023 V=14.0 ACC=20 DEC=20
MOVC C00024 V=14.0 ACC=20 DEC=20
MOVL C00025 V=10.0 ACC=20 DEC=20
MOVL C00026 V=10.0 ACC=20 DEC=20
MOVL C00027 V=10.0 ACC=20 DEC=20
MOVL C00028 V=10.0 ACC=20 DEC=20
MOVL C00029 V=10.0 ACC=20 DEC=20
MOVL C00030 V=10.0 ACC=20 DEC=20
MOVL C00031 V=10.0 ACC=20 DEC=20
MOVL C00032 V=10.0 ACC=20 DEC=20
MOVL C00033 V=10.0 ACC=20 DEC=20
MOVL C00034 V=10.0 ACC=20 DEC=20
MOVL C00035 V=10.0 ACC=20 DEC=20
MOVL C00036 V=10.0 ACC=20 DEC=20
MOVL C00037 V=10.0 ACC=20 DEC=20
MOVL C00038 V=10.0 ACC=20 DEC=20
MOVL C00039 V=10.0 ACC=20 DEC=20
MOVL C00040 V=10.0 ACC=20 DEC=20
MOVL C00041 V=10.0 ACC=20 DEC=20
MOVL C00042 V=10.0 ACC=20 DEC=20
MOVL C00043 V=10.0 ACC=20 DEC=20
MOVL C00044 V=10.0 ACC=20 DEC=20
ARCOF
TIMER T=60
MOVL C00045 V=11.0 ACC=20 DEC=20
*LAG2
MACRO1 MJ#(0) ARGF2
ARCON
MOVL C00046 V=10.0 ACC=20 DEC=20
MOVL C00047 V=10.0 ACC=20 DEC=20
MOVL C00048 V=10.0 ACC=20 DEC=20
MOVL C00049 V=10.0 ACC=20 DEC=20
MOVL C00050 V=10.0 ACC=20 DEC=20
MOVL C00051 V=10.0 ACC=20 DEC=20
MOVL C00052 V=10.0 ACC=20 DEC=20
MOVL C00053 V=10.0 ACC=20 DEC=20
MOVL C00054 V=10.0 ACC=20 DEC=20
MOVL C00055 V=10.0 ACC=20 DEC=20
MOVL C00056 V=10.0 ACC=20 DEC=20
MOVL C00057 V=10.0 ACC=20 DEC=20
MOVL C00058 V=10.0 ACC=20 DEC=20
MOVL C00059 V=10.0 ACC=20 DEC=20
MOVL C00060 V=10.0 ACC=20 DEC=20
MOVL C00061 V=10.0 ACC=20 DEC=20
MOVL C00062 V=10.0 ACC=20 DEC=20
MOVL C00063 V=10.0 ACC=20 DEC=20
MOVL C00064 V=10.0 ACC=20 DEC=20
MOVC C00065 V=14.0 ACC=20 DEC=20
MOVC C00066 V=14.0 ACC=20 DEC=20
MOVC C00067 V=14.0 ACC=20 DEC=20
MOVL C00068 V=10.0 ACC=20 DEC=20
MOVL C00069 V=10.0 ACC=20 DEC=20
MOVL C00070 V=10.0 ACC=20 DEC=20
MOVL C00071 V=10.0 ACC=20 DEC=20
MOVL C00072 V=10.0 ACC=20 DEC=20
MOVL C00073 V=10.0 ACC=20 DEC=20
MOVL C00074 V=10.0 ACC=20 DEC=20
MOVL C00075 V=10.0 ACC=20 DEC=20
MOVL C00076 V=10.0 ACC=20 DEC=20
MOVL C00077 V=10.0 ACC=20 DEC=20
MOVL C00078 V=10.0 ACC=20 DEC=20
MOVL C00079 V=10.0 ACC=20 DEC=20
MOVL C00080 V=10.0 ACC=20 DEC=20
MOVL C00081 V=10.0 ACC=20 DEC=20
MOVL C00082 V=10.0 ACC=20 DEC=20
MOVL C00083 V=10.0 ACC=20 DEC=20
MOVL C00084 V=10.0 ACC=20 DEC=20
MOVL C00085 V=10.0 ACC=20 DEC=20
MOVL C00086 V=10.0 ACC=20 DEC=20
MOVL C00087 V=10.0 ACC=20 DEC=20
ARCOF
TIMER T=60
MOVL C00088 V=11.0 ACC=20 DEC=20
*LAG3
MACRO1 MJ#(0) ARGF2
ARCON
MOVL C00089 V=10.0 ACC=20 DEC=20
MOVL C00090 V=10.0 ACC=20 DEC=20
MOVL C00091 V=10.0 ACC=20 DEC=20
MOVL C00092 V=10.0 ACC=20 DEC=20
MOVL C00093 V=10.0 ACC=20 DEC=20
MOVL C00094 V=10.0 ACC=20 DEC=20
MOVL C00095 V=10.0 ACC=20 DEC=20
MOVL C00096 V=10.0 ACC=20 DEC=20
MOVL C00097 V=10.0 ACC=20 DEC=20
MOVL C00098 V=10.0 ACC=20 DEC=20
MOVL C00099 V=10.0 ACC=20 DEC=20
MOVL C00100 V=10.0 ACC=20 DEC=20
MOVL C00101 V=10.0 ACC=20 DEC=20
MOVL C00102 V=10.0 ACC=20 DEC=20
MOVL C00103 V=10.0 ACC=20 DEC=20
MOVL C00104 V=10.0 ACC=20 DEC=20
MOVL C00105 V=10.0 ACC=20 DEC=20
MOVL C00106 V=10.0 ACC=20 DEC=20
MOVL C00107 V=10.0 ACC=20 DEC=20
MOVC C00108 V=14.0 ACC=20 DEC=20
MOVC C00109 V=14.0 ACC=20 DEC=20
MOVC C00110 V=14.0 ACC=20 DEC=20
MOVL C00111 V=10.0 ACC=20 DEC=20
MOVL C00112 V=10.0 ACC=20 DEC=20
MOVL C00113 V=10.0 ACC=20 DEC=20
MOVL C00114 V=10.0 ACC=20 DEC=20
MOVL C00115 V=10.0 ACC=20 DEC=20
MOVL C00116 V=10.0 ACC=20 DEC=20
MOVL C00117 V=10.0 ACC=20 DEC=20
MOVL C00118 V=10.0 ACC=20 DEC=20
MOVL C00119 V=10.0 ACC=20 DEC=20
MOVL C00120 V=10.0 ACC=20 DEC=20
MOVL C00121 V=10.0 ACC=20 DEC=20
MOVL C00122 V=10.0 ACC=20 DEC=20
MOVL C00123 V=10.0 ACC=20 DEC=20
MOVL C00124 V=10.0 ACC=20 DEC=20
MOVL C00125 V=10.0 ACC=20 DEC=20
MOVL C00126 V=10.0 ACC=20 DEC=20
MOVL C00127 V=10.0 ACC=20 DEC=20
MOVL C00128 V=10.0 ACC=20 DEC=20
MOVL C00129 V=10.0 ACC=20 DEC=20
MOVL C00130 V=10.0 ACC=20 DEC=20
ARCOF
TIMER T=60
MOVL C00131 V=11.0 ACC=20 DEC=20
*LAG4
MACRO1 MJ#(0) ARGF2
ARCON
MOVL C00132 V=10.0 ACC=20 DEC=20
MOVL C00133 V=10.0 ACC=20 DEC=20
MOVL C00134 V=10.0 ACC=20 DEC=20
MOVL C00135 V=10.0 ACC=20 DEC=20
MOVL C00136 V=10.0 ACC=20 DEC=20
MOVL C00137 V=10.0 ACC=20 DEC=20
MOVL C00138 V=10.0 ACC=20 DEC=20
MOVL C00139 V=10.0 ACC=20 DEC=20
MOVL C00140 V=10.0 ACC=20 DEC=20
MOVL C00141 V=10.0 ACC=20 DEC=20
MOVL C00142 V=10.0 ACC=20 DEC=20
MOVL C00143 V=10.0 ACC=20 DEC=20
MOVL C00144 V=10.0 ACC=20 DEC=20
MOVL C00145 V=10.0 ACC=20 DEC=20
MOVL C00146 V=10.0 ACC=20 DEC=20
MOVL C00147 V=10.0 ACC=20 DEC=20
MOVL C00148 V=10.0 ACC=20 DEC=20
MOVL C00149 V=10.0 ACC=20 DEC=20
MOVL C00150 V=10.0 ACC=20 DEC=20
MOVC C00151 V=14.0 ACC=20 DEC=20
MOVC C00152 V=14.0 ACC=20 DEC=20
MOVC C00153 V=14.0 ACC=20 DEC=20
MOVL C00154 V=10.0 ACC=20 DEC=20
MOVL C00155 V=10.0 ACC=20 DEC=20
MOVL C00156 V=10.0 ACC=20 DEC=20
MOVL C00157 V=10.0 ACC=20 DEC=20
MOVL C00158 V=10.0 ACC=20 DEC=20
MOVL C00159 V=10.0 ACC=20 DEC=20
MOVL C00160 V=10.0 ACC=20 DEC=20
MOVL C00161 V=10.0 ACC=20 DEC=20
MOVL C00162 V=10.0 ACC=20 DEC=20
MOVL C00163 V=10.0 ACC=20 DEC=20
MOVL C00164 V=10.0 ACC=20 DEC=20
MOVL C00165 V=10.0 ACC=20 DEC=20
MOVL C00166 V=10.0 ACC=20 DEC=20
MOVL C00167 V=10.0 ACC=20 DEC=20
MOVL C00168 V=10.0 ACC=20 DEC=20
MOVL C00169 V=10.0 ACC=20 DEC=20
MOVL C00170 V=10.0 ACC=20 DEC=20
MOVL C00171 V=10.0 ACC=20 DEC=20
MOVL C00172 V=10.0 ACC=20 DEC=20
MOVL C00173 V=10.0 ACC=20 DEC=20
ARCOF
TIMER T=60
MOVL C00174 V=11.0 ACC=20 DEC=20
*LAG5
MACRO1 MJ#(0) ARGF2
ARCON
MOVL C00175 V=10.0 ACC=20 DEC=20
MOVL C00176 V=10.0 ACC=20 DEC=20
MOVL C00177 V=10.0 ACC=20 DEC=20
MOVL C00178 V=10.0 ACC=20 DEC=20
MOVL C00179 V=10.0 ACC=20 DEC=20
MOVL C00180 V=10.0 ACC=20 DEC=20
MOVL C00181 V=10.0 ACC=20 DEC=20
MOVL C00182 V=10.0 ACC=20 DEC=20
MOVL C00183 V=10.0 ACC=20 DEC=20
MOVL C00184 V=10.0 ACC=20 DEC=20
MOVL C00185 V=10.0 ACC=20 DEC=20
MOVL C00186 V=10.0 ACC=20 DEC=20
MOVL C00187 V=10.0 ACC=20 DEC=20
MOVL C00188 V=10.0 ACC=20 DEC=20
MOVL C00189 V=10.0 ACC=20 DEC=20
MOVL C00190 V=10.0 ACC=20 DEC=20
MOVL C00191 V=10.0 ACC=20 DEC=20
MOVL C00192 V=10.0 ACC=20 DEC=20
MOVL C00193 V=10.0 ACC=20 DEC=20
MOVC C00194 V=14.0 ACC=20 DEC=20
MOVC C00195 V=14.0 ACC=20 DEC=20
MOVC C00196 V=14.0 ACC=20 DEC=20
MOVL C00197 V=10.0 ACC=20 DEC=20
MOVL C00198 V=10.0 ACC=20 DEC=20
MOVL C00199 V=10.0 ACC=20 DEC=20
MOVL C00200 V=10.0 ACC=20 DEC=20
MOVL C00201 V=10.0 ACC=20 DEC=20
MOVL C00202 V=10.0 ACC=20 DEC=20
MOVL C00203 V=10.0 ACC=20 DEC=20
MOVL C00204 V=10.0 ACC=20 DEC=20
MOVL C00205 V=10.0 ACC=20 DEC=20
MOVL C00206 V=10.0 ACC=20 DEC=20
MOVL C00207 V=10.0 ACC=20 DEC=20
MOVL C00208 V=10.0 ACC=20 DEC=20
MOVL C00209 V=10.0 ACC=20 DEC=20
MOVL C00210 V=10.0 ACC=20 DEC=20
MOVL C00211 V=10.0 ACC=20 DEC=20
MOVL C00212 V=10.0 ACC=20 DEC=20
MOVL C00213 V=10.0 ACC=20 DEC=20
MOVL C00214 V=10.0 ACC=20 DEC=20
MOVL C00215 V=10.0 ACC=20 DEC=20
MOVL C00216 V=10.0 ACC=20 DEC=20
ARCOF
TIMER T=60
MOVL C00217 V=11.0 ACC=20 DEC=20
*LAG6
MACRO1 MJ#(0) ARGF2
ARCON
MOVL C00218 V=10.0 ACC=20 DEC=20
MOVL C00219 V=10.0 ACC=20 DEC=20
MOVL C00220 V=10.0 ACC=20 DEC=20
MOVL C00221 V=10.0 ACC=20 DEC=20
MOVL C00222 V=10.0 ACC=20 DEC=20
MOVL C00223 V=10.0 ACC=20 DEC=20
MOVL C00224 V=10.0 ACC=20 DEC=20
MOVL C00225 V=10.0 ACC=20 DEC=20
MOVL C00226 V=10.0 ACC=20 DEC=20
MOVL C00227 V=10.0 ACC=20 DEC=20
MOVL C00228 V=10.0 ACC=20 DEC=20
MOVL C00229 V=10.0 ACC=20 DEC=20
MOVL C00230 V=10.0 ACC=20 DEC=20
MOVL C00231 V=10.0 ACC=20 DEC=20
MOVL C00232 V=10.0 ACC=20 DEC=20
MOVL C00233 V=10.0 ACC=20 DEC=20
MOVL C00234 V=10.0 ACC=20 DEC=20
MOVL C00235 V=10.0 ACC=20 DEC=20
MOVL C00236 V=10.0 ACC=20 DEC=20
MOVC C00237 V=14.0 ACC=20 DEC=20
MOVC C00238 V=14.0 ACC=20 DEC=20
MOVC C00239 V=14.0 ACC=20 DEC=20
MOVL C00240 V=10.0 ACC=20 DEC=20
MOVL C00241 V=10.0 ACC=20 DEC=20
MOVL C00242 V=10.0 ACC=20 DEC=20
MOVL C00243 V=10.0 ACC=20 DEC=20
MOVL C00244 V=10.0 ACC=20 DEC=20
MOVL C00245 V=10.0 ACC=20 DEC=20
MOVL C00246 V=10.0 ACC=20 DEC=20
MOVL C00247 V=10.0 ACC=20 DEC=20
MOVL C00248 V=10.0 ACC=20 DEC=20
MOVL C00249 V=10.0 ACC=20 DEC=20
MOVL C00250 V=10.0 ACC=20 DEC=20
MOVL C00251 V=10.0 ACC=20 DEC=20
MOVL C00252 V=10.0 ACC=20 DEC=20
MOVL C00253 V=10.0 ACC=20 DEC=20
MOVL C00254 V=10.0 ACC=20 DEC=20
MOVL C00255 V=10.0 ACC=20 DEC=20
MOVL C00256 V=10.0 ACC=20 DEC=20
MOVL C00257 V=10.0 ACC=20 DEC=20
MOVL C00258 V=10.0 ACC=20 DEC=20
MOVL C00259 V=10.0 ACC=20 DEC=20
ARCOF
TIMER T=60
MOVL C00260 V=11.0 ACC=20 DEC=20
*LAG7
MACRO1 MJ#(0) ARGF2
ARCON
MOVL C00261 V=10.0 ACC=20 DEC=20
MOVL C00262 V=10.0 ACC=20 DEC=20
MOVL C00263 V=10.0 ACC=20 DEC=20
MOVL C00264 V=10.0 ACC=20 DEC=20
MOVL C00265 V=10.0 ACC=20 DEC=20
MOVL C00266 V=10.0 ACC=20 DEC=20
MOVL C00267 V=10.0 ACC=20 DEC=20
MOVL C00268 V=10.0 ACC=20 DEC=20
MOVL C00269 V=10.0 ACC=20 DEC=20
MOVL C00270 V=10.0 ACC=20 DEC=20
MOVL C00271 V=10.0 ACC=20 DEC=20
MOVL C00272 V=10.0 ACC=20 DEC=20
MOVL C00273 V=10.0 ACC=20 DEC=20
MOVL C00274 V=10.0 ACC=20 DEC=20
MOVL C00275 V=10.0 ACC=20 DEC=20
MOVL C00276 V=10.0 ACC=20 DEC=20
MOVL C00277 V=10.0 ACC=20 DEC=20
MOVL C00278 V=10.0 ACC=20 DEC=20
MOVL C00279 V=10.0 ACC=20 DEC=20
MOVC C00280 V=14.0 ACC=20 DEC=20
MOVC C00281 V=14.0 ACC=20 DEC=20
MOVC C00282 V=14.0 ACC=20 DEC=20
MOVL C00283 V=10.0 ACC=20 DEC=20
MOVL C00284 V=10.0 ACC=20 DEC=20
MOVL C00285 V=10.0 ACC=20 DEC=20
MOVL C00286 V=10.0 ACC=20 DEC=20
MOVL C00287 V=10.0 ACC=20 DEC=20
MOVL C00288 V=10.0 ACC=20 DEC=20
MOVL C00289 V=10.0 ACC=20 DEC=20
MOVL C00290 V=10.0 ACC=20 DEC=20
MOVL C00291 V=10.0 ACC=20 DEC=20
MOVL C00292 V=10.0 ACC=20 DEC=20
MOVL C00293 V=10.0 ACC=20 DEC=20
MOVL C00294 V=10.0 ACC=20 DEC=20
MOVL C00295 V=10.0 ACC=20 DEC=20
MOVL C00296 V=10.0 ACC=20 DEC=20
MOVL C00297 V=10.0 ACC=20 DEC=20
MOVL C00298 V=10.0 ACC=20 DEC=20
MOVL C00299 V=10.0 ACC=20 DEC=20
MOVL C00300 V=10.0 ACC=20 DEC=20
MOVL C00301 V=10.0 ACC=20 DEC=20
MOVL C00302 V=10.0 ACC=20 DEC=20
ARCOF
TIMER T=60
MOVL C00303 V=11.0 ACC=20 DEC=20
*LAG8
MACRO1 MJ#(0) ARGF2
ARCON
MOVL C00304 V=10.0 ACC=20 DEC=20
MOVL C00305 V=10.0 ACC=20 DEC=20
MOVL C00306 V=10.0 ACC=20 DEC=20
MOVL C00307 V=10.0 ACC=20 DEC=20
MOVL C00308 V=10.0 ACC=20 DEC=20
MOVL C00309 V=10.0 ACC=20 DEC=20
MOVL C00310 V=10.0 ACC=20 DEC=20
MOVL C00311 V=10.0 ACC=20 DEC=20
MOVL C00312 V=10.0 ACC=20 DEC=20
MOVL C00313 V=10.0 ACC=20 DEC=20
MOVL C00314 V=10.0 ACC=20 DEC=20
MOVL C00315 V=10.0 ACC=20 DEC=20
MOVL C00316 V=10.0 ACC=20 DEC=20
MOVL C00317 V=10.0 ACC=20 DEC=20
MOVL C00318 V=10.0 ACC=20 DEC=20
MOVL C00319 V=10.0 ACC=20 DEC=20
MOVL C00320 V=10.0 ACC=20 DEC=20
MOVL C00321 V=10.0 ACC=20 DEC=20
MOVL C00322 V=10.0 ACC=20 DEC=20
MOVC C00323 V=14.0 ACC=20 DEC=20
MOVC C00324 V=14.0 ACC=20 DEC=20
MOVC C00325 V=14.0 ACC=20 DEC=20
MOVL C00326 V=10.0 ACC=20 DEC=20
MOVL C00327 V=10.0 ACC=20 DEC=20
MOVL C00328 V=10.0 ACC=20 DEC=20
MOVL C00329 V=10.0 ACC=20 DEC=20
MOVL C00330 V=10.0 ACC=20 DEC=20
MOVL C00331 V=10.0 ACC=20 DEC=20
MOVL C00332 V=10.0 ACC=20 DEC=20
MOVL C00333 V=10.0 ACC=20 DEC=20
MOVL C00334 V=10.0 ACC=20 DEC=20
MOVL C00335 V=10.0 ACC=20 DEC=20
MOVL C00336 V=10.0 ACC=20 DEC=20
MOVL C00337 V=10.0 ACC=20 DEC=20
MOVL C00338 V=10.0 ACC=20 DEC=20
MOVL C00339 V=10.0 ACC=20 DEC=20
MOVL C00340 V=10.0 ACC=20 DEC=20
MOVL C00341 V=10.0 ACC=20 DEC=20
MOVL C00342 V=10.0 ACC=20 DEC=20
MOVL C00343 V=10.0 ACC=20 DEC=20
MOVL C00344 V=10.0 ACC=20 DEC=20
MOVL C00345 V=10.0 ACC=20 DEC=20
ARCOF
TIMER T=60
MOVL C00346 V=11.0 ACC=20 DEC=20
*LAG9
MACRO1 MJ#(0) ARGF2
ARCON
MOVL C00347 V=10.0 ACC=20 DEC=20
MOVL C00348 V=10.0 ACC=20 DEC=20
MOVL C00349 V=10.0 ACC=20 DEC=20
MOVL C00350 V=10.0 ACC=20 DEC=20
MOVL C00351 V=10.0 ACC=20 DEC=20
MOVL C00352 V=10.0 ACC=20 DEC=20
MOVL C00353 V=10.0 ACC=20 DEC=20
MOVL C00354 V=10.0 ACC=20 DEC=20
MOVL C00355 V=10.0 ACC=20 DEC=20
MOVL C00356 V=10.0 ACC=20 DEC=20
MOVL C00357 V=10.0 ACC=20 DEC=20
MOVL C00358 V=10.0 ACC=20 DEC=20
MOVL C00359 V=10.0 ACC=20 DEC=20
MOVL C00360 V=10.0 ACC=20 DEC=20
MOVL C00361 V=10.0 ACC=20 DEC=20
MOVL C00362 V=10.0 ACC=20 DEC=20
MOVL C00363 V=10.0 ACC=20 DEC=20
MOVL C00364 V=10.0 ACC=20 DEC=20
MOVL C00365 V=10.0 ACC=20 DEC=20
MOVC C00366 V=14.0 ACC=20 DEC=20
MOVC C00367 V=14.0 ACC=20 DEC=20
MOVC C00368 V=14.0 ACC=20 DEC=20
MOVL C00369 V=10.0 ACC=20 DEC=20
MOVL C00370 V=10.0 ACC=20 DEC=20
MOVL C00371 V=10.0 ACC=20 DEC=20
MOVL C00372 V=10.0 ACC=20 DEC=20
MOVL C00373 V=10.0 ACC=20 DEC=20
MOVL C00374 V=10.0 ACC=20 DEC=20
MOVL C00375 V=10.0 ACC=20 DEC=20
MOVL C00376 V=10.0 ACC=20 DEC=20
MOVL C00377 V=10.0 ACC=20 DEC=20
MOVL C00378 V=10.0 ACC=20 DEC=20
MOVL C00379 V=10.0 ACC=20 DEC=20
MOVL C00380 V=10.0 ACC=20 DEC=20
MOVL C00381 V=10.0 ACC=20 DEC=20
MOVL C00382 V=10.0 ACC=20 DEC=20
MOVL C00383 V=10.0 ACC=20 DEC=20
MOVL C00384 V=10.0 ACC=20 DEC=20
MOVL C00385 V=10.0 ACC=20 DEC=20
MOVL C00386 V=10.0 ACC=20 DEC=20
MOVL C00387 V=10.0 ACC=20 DEC=20
MOVL C00388 V=10.0 ACC=20 DEC=20
ARCOF
TIMER T=60
MOVL C00389 V=11.0 ACC=20 DEC=20
*LAG10
MACRO1 MJ#(0) ARGF2
ARCON
MOVL C00390 V=10.0 ACC=20 DEC=20
MOVL C00391 V=10.0 ACC=20 DEC=20
MOVL C00392 V=10.0 ACC=20 DEC=20
MOVL C00393 V=10.0 ACC=20 DEC=20
MOVL C00394 V=10.0 ACC=20 DEC=20
MOVL C00395 V=10.0 ACC=20 DEC=20
MOVL C00396 V=10.0 ACC=20 DEC=20
MOVL C00397 V=10.0 ACC=20 DEC=20
MOVL C00398 V=10.0 ACC=20 DEC=20
MOVL C00399 V=10.0 ACC=20 DEC=20
MOVL C00400 V=10.0 ACC=20 DEC=20
MOVL C00401 V=10.0 ACC=20 DEC=20
MOVL C00402 V=10.0 ACC=20 DEC=20
MOVL C00403 V=10.0 ACC=20 DEC=20
MOVL C00404 V=10.0 ACC=20 DEC=20
MOVL C00405 V=10.0 ACC=20 DEC=20
MOVL C00406 V=10.0 ACC=20 DEC=20
MOVL C00407 V=10.0 ACC=20 DEC=20
MOVL C00408 V=10.0 ACC=20 DEC=20
MOVC C00409 V=14.0 ACC=20 DEC=20
MOVC C00410 V=14.0 ACC=20 DEC=20
MOVC C00411 V=14.0 ACC=20 DEC=20
MOVL C00412 V=10.0 ACC=20 DEC=20
MOVL C00413 V=10.0 ACC=20 DEC=20
MOVL C00414 V=10.0 ACC=20 DEC=20
MOVL C00415 V=10.0 ACC=20 DEC=20
MOVL C00416 V=10.0 ACC=20 DEC=20
MOVL C00417 V=10.0 ACC=20 DEC=20
MOVL C00418 V=10.0 ACC=20 DEC=20
MOVL C00419 V=10.0 ACC=20 DEC=20
MOVL C00420 V=10.0 ACC=20 DEC=20
MOVL C00421 V=10.0 ACC=20 DEC=20
MOVL C00422 V=10.0 ACC=20 DEC=20
MOVL C00423 V=10.0 ACC=20 DEC=20
MOVL C00424 V=10.0 ACC=20 DEC=20
MOVL C00425 V=10.0 ACC=20 DEC=20
MOVL C00426 V=10.0 ACC=20 DEC=20
MOVL C00427 V=10.0 ACC=20 DEC=20
MOVL C00428 V=10.0 ACC=20 DEC=20
MOVL C00429 V=10.0 ACC=20 DEC=20
MOVL C00430 V=10.0 ACC=20 DEC=20
MOVL C00431 V=10.0 ACC=20 DEC=20
ARCOF
TIMER T=60
MOVL C00432 V=11.0 ACC=20 DEC=20
*LAG11
MACRO1 MJ#(0) ARGF2
ARCON
MOVL C00433 V=10.0 ACC=20 DEC=20
MOVL C00434 V=10.0 ACC=20 DEC=20
MOVL C00435 V=10.0 ACC=20 DEC=20
MOVL C00436 V=10.0 ACC=20 DEC=20
MOVL C00437 V=10.0 ACC=20 DEC=20
MOVL C00438 V=10.0 ACC=20 DEC=20
MOVL C00439 V=10.0 ACC=20 DEC=20
MOVL C00440 V=10.0 ACC=20 DEC=20
MOVL C00441 V=10.0 ACC=20 DEC=20
MOVL C00442 V=10.0 ACC=20 DEC=20
MOVL C00443 V=10.0 ACC=20 DEC=20
MOVL C00444 V=10.0 ACC=20 DEC=20
MOVL C00445 V=10.0 ACC=20 DEC=20
MOVL C00446 V=10.0 ACC=20 DEC=20
MOVL C00447 V=10.0 ACC=20 DEC=20
MOVL C00448 V=10.0 ACC=20 DEC=20
MOVL C00449 V=10.0 ACC=20 DEC=20
MOVL C00450 V=10.0 ACC=20 DEC=20
MOVL C00451 V=10.0 ACC=20 DEC=20
MOVC C00452 V=14.0 ACC=20 DEC=20
MOVC C00453 V=14.0 ACC=20 DEC=20
MOVC C00454 V=14.0 ACC=20 DEC=20
MOVL C00455 V=10.0 ACC=20 DEC=20
MOVL C00456 V=10.0 ACC=20 DEC=20
MOVL C00457 V=10.0 ACC=20 DEC=20
MOVL C00458 V=10.0 ACC=20 DEC=20
MOVL C00459 V=10.0 ACC=20 DEC=20
MOVL C00460 V=10.0 ACC=20 DEC=20
MOVL C00461 V=10.0 ACC=20 DEC=20
MOVL C00462 V=10.0 ACC=20 DEC=20
MOVL C00463 V=10.0 ACC=20 DEC=20
MOVL C00464 V=10.0 ACC=20 DEC=20
MOVL C00465 V=10.0 ACC=20 DEC=20
MOVL C00466 V=10.0 ACC=20 DEC=20
MOVL C00467 V=10.0 ACC=20 DEC=20
MOVL C00468 V=10.0 ACC=20 DEC=20
MOVL C00469 V=10.0 ACC=20 DEC=20
MOVL C00470 V=10.0 ACC=20 DEC=20
MOVL C00471 V=10.0 ACC=20 DEC=20
MOVL C00472 V=10.0 ACC=20 DEC=20
MOVL C00473 V=10.0 ACC=20 DEC=20
MOVL C00474 V=10.0 ACC=20 DEC=20
ARCOF
TIMER T=60
MOVL C00475 V=11.0 ACC=20 DEC=20
*LAG12
MACRO1 MJ#(0) ARGF2
ARCON
MOVL C00476 V=10.0 ACC=20 DEC=20
MOVL C00477 V=10.0 ACC=20 DEC=20
MOVL C00478 V=10.0 ACC=20 DEC=20
MOVL C00479 V=10.0 ACC=20 DEC=20
MOVL C00480 V=10.0 ACC=20 DEC=20
MOVL C00481 V=10.0 ACC=20 DEC=20
MOVL C00482 V=10.0 ACC=20 DEC=20
MOVL C00483 V=10.0 ACC=20 DEC=20
MOVL C00484 V=10.0 ACC=20 DEC=20
MOVL C00485 V=10.0 ACC=20 DEC=20
MOVL C00486 V=10.0 ACC=20 DEC=20
MOVL C00487 V=10.0 ACC=20 DEC=20
MOVL C00488 V=10.0 ACC=20 DEC=20
MOVL C00489 V=10.0 ACC=20 DEC=20
MOVL C00490 V=10.0 ACC=20 DEC=20
MOVL C00491 V=10.0 ACC=20 DEC=20
MOVL C00492 V=10.0 ACC=20 DEC=20
MOVL C00493 V=10.0 ACC=20 DEC=20
MOVL C00494 V=10.0 ACC=20 DEC=20
MOVC C00495 V=14.0 ACC=20 DEC=20
MOVC C00496 V=14.0 ACC=20 DEC=20
MOVC C00497 V=14.0 ACC=20 DEC=20
MOVL C00498 V=10.0 ACC=20 DEC=20
MOVL C00499 V=10.0 ACC=20 DEC=20
MOVL C00500 V=10.0 ACC=20 DEC=20
MOVL C00501 V=10.0 ACC=20 DEC=20
MOVL C00502 V=10.0 ACC=20 DEC=20
MOVL C00503 V=10.0 ACC=20 DEC=20
MOVL C00504 V=10.0 ACC=20 DEC=20
MOVL C00505 V=10.0 ACC=20 DEC=20
MOVL C00506 V=10.0 ACC=20 DEC=20
MOVL C00507 V=10.0 ACC=20 DEC=20
MOVL C00508 V=10.0 ACC=20 DEC=20
MOVL C00509 V=10.0 ACC=20 DEC=20
MOVL C00510 V=10.0 ACC=20 DEC=20
MOVL C00511 V=10.0 ACC=20 DEC=20
MOVL C00512 V=10.0 ACC=20 DEC=20
MOVL C00513 V=10.0 ACC=20 DEC=20
MOVL C00514 V=10.0 ACC=20 DEC=20
MOVL C00515 V=10.0 ACC=20 DEC=20
MOVL C00516 V=10.0 ACC=20 DEC=20
MOVL C00517 V=10.0 ACC=20 DEC=20
ARCOF
TIMER T=60
MOVL C00518 V=11.0 ACC=20 DEC=20
*LAG13
MACRO1 MJ#(0) ARGF2
ARCON
MOVL C00519 V=10.0 ACC=20 DEC=20
MOVL C00520 V=10.0 ACC=20 DEC=20
MOVL C00521 V=10.0 ACC=20 DEC=20
MOVL C00522 V=10.0 ACC=20 DEC=20
MOVL C00523 V=10.0 ACC=20 DEC=20
MOVL C00524 V=10.0 ACC=20 DEC=20
MOVL C00525 V=10.0 ACC=20 DEC=20
MOVL C00526 V=10.0 ACC=20 DEC=20
MOVL C00527 V=10.0 ACC=20 DEC=20
MOVL C00528 V=10.0 ACC=20 DEC=20
MOVL C00529 V=10.0 ACC=20 DEC=20
MOVL C00530 V=10.0 ACC=20 DEC=20
MOVL C00531 V=10.0 ACC=20 DEC=20
MOVL C00532 V=10.0 ACC=20 DEC=20
MOVL C00533 V=10.0 ACC=20 DEC=20
MOVL C00534 V=10.0 ACC=20 DEC=20
MOVL C00535 V=10.0 ACC=20 DEC=20
MOVL C00536 V=10.0 ACC=20 DEC=20
MOVL C00537 V=10.0 ACC=20 DEC=20
MOVC C00538 V=14.0 ACC=20 DEC=20
MOVC C00539 V=14.0 ACC=20 DEC=20
MOVC C00540 V=14.0 ACC=20 DEC=20
MOVL C00541 V=10.0 ACC=20 DEC=20
MOVL C00542 V=10.0 ACC=20 DEC=20
MOVL C00543 V=10.0 ACC=20 DEC=20
MOVL C00544 V=10.0 ACC=20 DEC=20
MOVL C00545 V=10.0 ACC=20 DEC=20
MOVL C00546 V=10.0 ACC=20 DEC=20
MOVL C00547 V=10.0 ACC=20 DEC=20
MOVL C00548 V=10.0 ACC=20 DEC=20
MOVL C00549 V=10.0 ACC=20 DEC=20
MOVL C00550 V=10.0 ACC=20 DEC=20
MOVL C00551 V=10.0 ACC=20 DEC=20
MOVL C00552 V=10.0 ACC=20 DEC=20
MOVL C00553 V=10.0 ACC=20 DEC=20
MOVL C00554 V=10.0 ACC=20 DEC=20
MOVL C00555 V=10.0 ACC=20 DEC=20
MOVL C00556 V=10.0 ACC=20 DEC=20
MOVL C00557 V=10.0 ACC=20 DEC=20
MOVL C00558 V=10.0 ACC=20 DEC=20
MOVL C00559 V=10.0 ACC=20 DEC=20
MOVL C00560 V=10.0 ACC=20 DEC=20
ARCOF
TIMER T=60
MOVL C00561 V=11.0 ACC=20 DEC=20
*LAG14
MACRO1 MJ#(0) ARGF2
ARCON
MOVL C00562 V=10.0 ACC=20 DEC=20
MOVL C00563 V=10.0 ACC=20 DEC=20
MOVL C00564 V=10.0 ACC=20 DEC=20
MOVL C00565 V=10.0 ACC=20 DEC=20
MOVL C00566 V=10.0 ACC=20 DEC=20
MOVL C00567 V=10.0 ACC=20 DEC=20
MOVL C00568 V=10.0 ACC=20 DEC=20
MOVL C00569 V=10.0 ACC=20 DEC=20
MOVL C00570 V=10.0 ACC=20 DEC=20
MOVL C00571 V=10.0 ACC=20 DEC=20
MOVL C00572 V=10.0 ACC=20 DEC=20
MOVL C00573 V=10.0 ACC=20 DEC=20
MOVL C00574 V=10.0 ACC=20 DEC=20
MOVL C00575 V=10.0 ACC=20 DEC=20
MOVL C00576 V=10.0 ACC=20 DEC=20
MOVL C00577 V=10.0 ACC=20 DEC=20
MOVL C00578 V=10.0 ACC=20 DEC=20
MOVL C00579 V=10.0 ACC=20 DEC=20
MOVL C00580 V=10.0 ACC=20 DEC=20
MOVC C00581 V=14.0 ACC=20 DEC=20
MOVC C00582 V=14.0 ACC=20 DEC=20
MOVC C00583 V=14.0 ACC=20 DEC=20
MOVL C00584 V=10.0 ACC=20 DEC=20
MOVL C00585 V=10.0 ACC=20 DEC=20
MOVL C00586 V=10.0 ACC=20 DEC=20
MOVL C00587 V=10.0 ACC=20 DEC=20
MOVL C00588 V=10.0 ACC=20 DEC=20
MOVL C00589 V=10.0 ACC=20 DEC=20
MOVL C00590 V=10.0 ACC=20 DEC=20
MOVL C00591 V=10.0 ACC=20 DEC=20
MOVL C00592 V=10.0 ACC=20 DEC=20
MOVL C00593 V=10.0 ACC=20 DEC=20
MOVL C00594 V=10.0 ACC=20 DEC=20
MOVL C00595 V=10.0 ACC=20 DEC=20
MOVL C00596 V=10.0 ACC=20 DEC=20
MOVL C00597 V=10.0 ACC=20 DEC=20
MOVL C00598 V=10.0 ACC=20 DEC=20
MOVL C00599 V=10.0 ACC=20 DEC=20
MOVL C00600 V=10.0 ACC=20 DEC=20
MOVL C00601 V=10.0 ACC=20 DEC=20
MOVL C00602 V=10.0 ACC=20 DEC=20
MOVL C00603 V=10.0 ACC=20 DEC=20
ARCOF
TIMER T=60
MOVL C00604 V=11.0 ACC=20 DEC=20
*LAG15
MACRO1 MJ#(0) ARGF2
ARCON
MOVL C00605 V=10.0 ACC=20 DEC=20
MOVL C00606 V=10.0 ACC=20 DEC=20
MOVL C00607 V=10.0 ACC=20 DEC=20
MOVL C00608 V=10.0 ACC=20 DEC=20
MOVL C00609 V=10.0 ACC=20 DEC=20
MOVL C00610 V=10.0 ACC=20 DEC=20
MOVL C00611 V=10.0 ACC=20 DEC=20
MOVL C00612 V=10.0 ACC=20 DEC=20
MOVL C00613 V=10.0 ACC=20 DEC=20
MOVL C00614 V=10.0 ACC=20 DEC=20
MOVL C00615 V=10.0 ACC=20 DEC=20
MOVL C00616 V=10.0 ACC=20 DEC=20
MOVL C00617 V=10.0 ACC=20 DEC=20
MOVL C00618 V=10.0 ACC=20 DEC=20
MOVL C00619 V=10.0 ACC=20 DEC=20
MOVL C00620 V=10.0 ACC=20 DEC=20
MOVL C00621 V=10.0 ACC=20 DEC=20
MOVL C00622 V=10.0 ACC=20 DEC=20
MOVL C00623 V=10.0 ACC=20 DEC=20
MOVC C00624 V=14.0 ACC=20 DEC=20
MOVC C00625 V=14.0 ACC=20 DEC=20
MOVC C00626 V=14.0 ACC=20 DEC=20
MOVL C00627 V=10.0 ACC=20 DEC=20
MOVL C00628 V=10.0 ACC=20 DEC=20
MOVL C00629 V=10.0 ACC=20 DEC=20
MOVL C00630 V=10.0 ACC=20 DEC=20
MOVL C00631 V=10.0 ACC=20 DEC=20
MOVL C00632 V=10.0 ACC=20 DEC=20
MOVL C00633 V=10.0 ACC=20 DEC=20
MOVL C00634 V=10.0 ACC=20 DEC=20
MOVL C00635 V=10.0 ACC=20 DEC=20
MOVL C00636 V=10.0 ACC=20 DEC=20
MOVL C00637 V=10.0 ACC=20 DEC=20
MOVL C00638 V=10.0 ACC=20 DEC=20
MOVL C00639 V=10.0 ACC=20 DEC=20
MOVL C00640 V=10.0 ACC=20 DEC=20
MOVL C00641 V=10.0 ACC=20 DEC=20
MOVL C00642 V=10.0 ACC=20 DEC=20
MOVL C00643 V=10.0 ACC=20 DEC=20
MOVL C00644 V=10.0 ACC=20 DEC=20
MOVL C00645 V=10.0 ACC=20 DEC=20
MOVL C00646 V=10.0 ACC=20 DEC=20
ARCOF
TIMER T=60
MOVL C00647 V=11.0 ACC=20 DEC=20
MOVJ C00648 VJ=0.78
END
